(* IEC 61131-3 sources: rusty/tests/lit/cfc/blocks/expression_pin, 2 files *)

(* ---- main.st ---- *)
FUNCTION main : DINT
    expression_pin();
    expression_pin();
    // CHECK: a = 4, b = 44
    printf('a = %d, b = %d$N', expression_pin.outA, expression_pin.outB);
END_FUNCTION

(* ---- counter.st ---- *)
FUNCTION_BLOCK counter
VAR_INPUT
    step : DINT;
END_VAR
VAR_OUTPUT
    total : DINT;
END_VAR
    total := total + step;
END_FUNCTION_BLOCK
